FUNCTION_BLOCK FB_REF_Laser
VAR_INPUT
    {attribute 'pytmc' := '
        pv: SHUTDOWN
        io: io
    '}
    bShutdown: BOOL;

    {attribute 'pytmc' := '
        pv: PCT
        io: io
    '}
    fLaserPercent: LREAL;

    fTermMax: LREAL := 200;
END_VAR
VAR
    iShutdownINT AT %Q*: INT;
    iLaserINT AT %Q*: INT;

    fbGetLasPercent: FB_AnalogInput;
    fbSetLasPercent: FB_AnalogOutput;
END_VAR

// Send 5V to suppress laser
IF bShutdown THEN
    iShutdownINT := LREAL_TO_INT(EXPT(2, 14));
ELSE
    iShutdownINT := 0;
END_IF

// Limit to 0-5V instead of 10V
fbSetLasPercent(
    fReal:=fLaserPercent,
    fSafeMax:=100,
    fSafeMin:=0,
    iTermBits:=15,
    fTermMax:=fTermMax,
    fTermMin:=0,
    iRaw=>iLaserInt);
fbGetLasPercent(
    iRaw:=iLaserInt,
    iTermBits:=15,
    fTermMax:=fTermMax,
    fTermMin:=0,
    fReal=>fLaserPercent);

END_FUNCTION_BLOCK

(* stored: Version 1.1.0.1
   POU FB_REF_Laser: Id {fe34aa45-49f5-4ca6-ae16-2db42771e34d}, SpecialFunc None *)
